(*
This is a top-level paragraph.

    This paragraph belongs to a first-level block quote.

    This is the second paragraph of the first-level block quote.

        This paragraph belongs to a second-level block quote.

Another top-level paragraph.

        This paragraph belongs to a second-level block quote.

    This paragraph belongs to a first-level block quote. The
    second-level block quote above is inside this first-level
    block quote.
*)

FUNCTION_BLOCK FB_Libdoc_BlockQuote
VAR_INPUT
    nVarA : INT;
    nVarB : INT;
END_VAR
VAR_OUTPUT
    nSum : INT;
END_VAR
VAR
END_VAR

END_FUNCTION_BLOCK

(* stored: Version 1.1.0.1, ProductVersion 3.1.4022.18
   POU FB_Libdoc_BlockQuote: Id {f16f8a72-abf4-4e11-b54c-928318ad3314}, SpecialFunc None *)
